(* IEC 61131-3 sources: SortJet_MasterSPS_Aufbau.fbsproj/09_Station/UnterStationsbausteine/Entwicklung, 3 files *)

(* ---- Geblaese_Motorstarter_FB_V01_00_00.fb.st ---- *)
(* METADATA
{
	"v3Meta": {
		"objectGuid": "dfcb45a0-2101-41d2-aaa7-f1a51c527b1b"
	}
}
*)
{attribute 'excludefrombuild'}
FUNCTION_BLOCK Geblaese_Motorstarter_FB_V01_00_00 EXTENDS Geblaese_Schuetz_FB_V01_00_00
VAR_INPUT

END_VAR
VAR_OUTPUT
END_VAR
VAR
END_VAR

//-------------------------------------------------------------------------------------------------
// MASTER AUFRUFEN
//-------------------------------------------------------------------------------------------------
SUPER^(BasisStationsParameter := BasisStationsParameter);
END_FUNCTION_BLOCK

(* ---- Hub_FB_Methode_V01_00_00.fb.st ---- *)
(* METADATA
{
	"v3Meta": {
		"objectGuid": "edcc4463-460d-49b8-9b6c-0b51cf9d081d"
	}
}
*)
{attribute 'excludefrombuild'}
FUNCTION_BLOCK Hub_FB_Methode_V01_00_00
VAR_INPUT

  // BOOLEAN
  bpAktivieren               : BOOL;
  bpStartHubAuf              : BOOL;
  bpStartHubAb               : BOOL;
  bpReset                    : BOOL;
  bpSensorEinlaufNachfolger  : BOOL;
  bpSensorAuslaufVorgaenger  : BOOL;
  bpSensorEinlauf            : BOOL;
  bpSensorAuslauf            : BOOL;

  // STRUCT
  stStationsNummern          : Station_ST;

// POINTER *)
//ppParameterBaustein        : REFERENCE TO Parameter_Hub; // Zeiger auf Parameterfeld

END_VAR
VAR_OUTPUT

  // BOOLEAN
  bpFehler        : BOOL;
  bpDone          : BOOL;
  bpResourceAktiv : BOOL;

  // WORD
  wpFehlerNr : Fehlerkonstanten_EN;

  // ENUM
  epHubStatus  : Hub_EN; // Status: Gibt die Aktuelle Position des Antriebs aus

END_VAR

VAR

  // BOOLEAN
  blErsterZyklus        : BOOL := TRUE;

  // TIMER
  tonlMaxWarteZeit                        : TON;
  tonlHubAntriebOK                        : TON;
  tonlMaximaleWartezeitAufReset           : TON;
  tonlFehlermeldungUnterdrueckenAntriebOK : TON;
  tonlReset                               : TON;

  // TRIGGER
  ftrigFehlerAmSteuerteil : F_TRIG;

  // STEPS
  steplHubAb    : Steps_TE;
  steplHubAuf   : Steps_TE;
  steplReset    : Steps_TE;

  Motorstarter : Motorstarter_FB_V01_00_00;

END_VAR

VAR
  // HARDWARE EINGÄNGE
  in_bSensorNichtUnten             AT%I* : BOOL;
  in_bSensorNichtOben              AT%I* : BOOL;
  in_bMotorstarter_OK              AT%I* : BOOL;
  in_bLSBremse_OK                  AT%I* : BOOL;
  in_bLS400V_OK                    AT%I* : BOOL;

  // HARDWARE AUSGÄNGE
  out_bHubAbSetzen                 AT%Q* : BOOL;
  out_bHubAufSetzen                AT%Q* : BOOL;
  out_bReset                       AT%Q* : BOOL;
  out_bBremseLoesen                AT%Q* : BOOL;

END_VAR

VAR CONSTANT

  // TIME
  ZEITWERT_RESOURCE_AKTIV_AUSSCHALT_VERZOEGERN : TIME := T#25ms;

END_VAR

//-------------------------------------------------------------------------------------------------
// BAUSTEIN: INITIALISIERUNG
//-------------------------------------------------------------------------------------------------
IF ( blErsterZyklus ) THEN
  blErsterZyklus := FALSE;

  (* Hinweis:
     - Timer initialisieren
  *)
  tonlHubAntriebOK(IN:=TRUE);
  tonlMaxWarteZeit(IN:=FALSE);
  tonlFehlermeldungUnterdrueckenAntriebOK( IN := FALSE );

END_IF

//-------------------------------------------------------------------------------------------------
// BAUSTEIN: AKTIONEN
//-------------------------------------------------------------------------------------------------
IF ( bpAktivieren ) THEN
  Motorstarter();

  IF bpReset THEN
    wpFehlerNr := cMELDUNG_NULL;
    bpFehler   := FALSE;
    Motorstarter.Reset();

  ELSIF bpFehler THEN
    ;

  ELSIF bpStartHubAuf THEN
    bpDone := Motorstarter.Linkslauf();

  ELSIF  bpStartHubAb THEN
    bpDone := Motorstarter.Rechtslauf();

  END_IF

  Ausgaenge();
  Meldungen();
  Timer();

ELSE

  bpDone   := TRUE;
  bpFehler := FALSE;

  IF (bpStartHubAb AND NOT bpStartHubAuf) THEN
    epHubStatus := eHub_Unten;
  ELSIF (bpStartHubAuf AND NOT bpStartHubAb) THEN
    epHubStatus := eHub_Oben;
  ELSIF (bpStartHubAb AND NOT bpStartHubAuf) THEN
    epHubStatus := eHub_Undefiniert;
  END_IF

END_IF
END_FUNCTION_BLOCK

(* ---- Motorstarter_FB_V01_00_00.fb.st ---- *)
(* METADATA
{
	"v3Meta": {
		"objectGuid": "7ae6aadb-d504-4a64-ae44-49a559d1f9ad"
	}
}
*)
{attribute 'excludefrombuild'}
FUNCTION_BLOCK Motorstarter_FB_V01_00_00
VAR_INPUT
  bpReset                    : BOOL;
  bpMotorstarterOK           : BOOL;
  bpSensorNotNockeLinkslauf  : BOOL;
  bpSensorNotNockeRechtslauf : BOOL;
END_VAR
VAR_OUTPUT
  bpFehler   : BOOL;
  bpdone     : BOOL;

  wpFehlerNr : Fehlerkonstanten_EN;

  // IO's
  out_bLinkslauf   : BOOL;
  out_bRechtslauf  : BOOL;
  out_Reset        : BOOL;
  out_BremseLoesen : BOOL;

END_VAR
VAR
  // BOOLEAN
  blErsterZyklus : BOOL := TRUE;

  // TIMER
  tonlFehlermeldungUnterdrueckenAntriebOK : TON;

END_VAR

(* Hinweis:
   - Um nicht beim Starten der Anlage in einem Fehler zustehen (HubAntrieb Fehler ist Zeitgesteuert),
     wird der Fehler erst nach einigen Sekunden nach dem ersten Durchlaufen dieses Bausteins ausgewertet
*)
tonlFehlermeldungUnterdrueckenAntriebOK( IN := NOT blErsterZyklus,
                                         PT := T#4s );

IF bpReset THEN
  bpdone := Reset();
ELSIF bpFehler THEN
  out_bLinkslauf  := FALSE;
  out_bRechtslauf := FALSE;
ELSE
  bpdone := FALSE;
END_IF

// Bremse lösen
out_BremseLoesen := out_bLinkslauf OR out_bRechtslauf;
END_FUNCTION_BLOCK
